// TIA Portal V21 export
// export: Created 2026-11-10T07:35:24.3181512Z, ExportSetting WithDefaults, DisplayName Totally Integrated Automation Portal, DisplayVersion V21 Update 3, DisplayName STEP 7 Professional, DisplayVersion V21 Update 3, DisplayName STEP 7 Safety, DisplayVersion V21, DisplayName Tech WebApplication, DisplayVersion V21, DisplayName WinCC Basic/Comfort/Advanced, DisplayVersion V21 Update 3, DisplayName WinCC Unified, DisplayVersion V21 Update 3
FUNCTION_BLOCK "FB_Lad_ex160"   // FB61, LAD
{ S7_Optimized_Access := 'TRUE' }
VERSION : 0.1
// stored: AutoNumber true, IsIECCheckEnabled false, IsRetainMemResEnabled false, MemoryReserve 100, SetENOAutomatically false, UDAEnableTagReadback false
   VAR_INPUT
      v_subnetid : Byte;
      v_rack : Word;
      v_slot : Word;
      v_subslot : Byte;
      v_subaddr : Word;
      v_ret_val : Int;
   END_VAR
   VAR_OUTPUT
      v_ioid : Byte;
      v_laddr : HW_MODULE;
   END_VAR
BEGIN

REGION Network 1: GADR_LGC - Determine hardware identifier from slot and offset in the user data address area
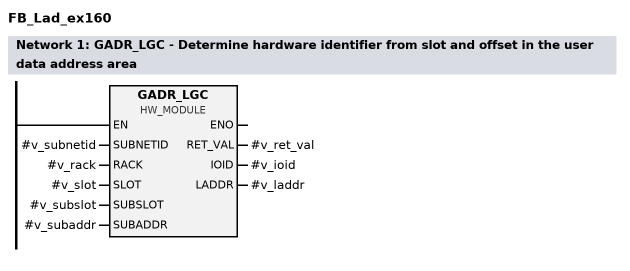
   RUNG wire#powerrail
      { S7_Templates := "laddr_type := HW_MODULE" } GADR_LGC(SUBNETID := #v_subnetid, RACK := #v_rack, SLOT := #v_slot, SUBSLOT := #v_subslot, SUBADDR := #v_subaddr, RET_VAL => #v_ret_val, IOID => #v_ioid, LADDR => #v_laddr)
   END_RUNG
   // the same network as SCL:
   #v_ret_val := GADR_LGC(SUBNETID := #v_subnetid,
                          RACK := #v_rack,
                          SLOT := #v_slot,
                          SUBSLOT := #v_subslot,
                          SUBADDR := #v_subaddr,
                          IOID => #v_ioid,
                          LADDR => #v_laddr);
END_REGION
END_FUNCTION_BLOCK
